Fanuc KAREL source: KA00115.KL

PROGRAM KA00115
%NOLOCKGROUP
VAR
  SRC: CONFIG
  DST: XYZWPREXT
BEGIN
  SRC.CFG_FLIP = TRUE
  DST = SRC
END KA00115
